(* PLC project AgentPLC, Beckhoff Automation GmbH TwinCAT PLC Control 3.5.21.61 *)
(* stored: creationDateTime 2026-11-03T10:24:45.563819, modificationDateTime 2026-11-03T10:24:45.5668157 *)

PROGRAM MAIN
VAR
	StartPB : BOOL;
	StopNC : BOOL;
	EStopHealthy : BOOL;
	PartSensor : BOOL;
	CountReset : BOOL;
	RunReq : BOOL;
	Horn : BOOL;
	Motor : BOOL;
	BatchLamp : BOOL;
	StartDelay : TON;
	BatchCounter : CTU;
END_VAR

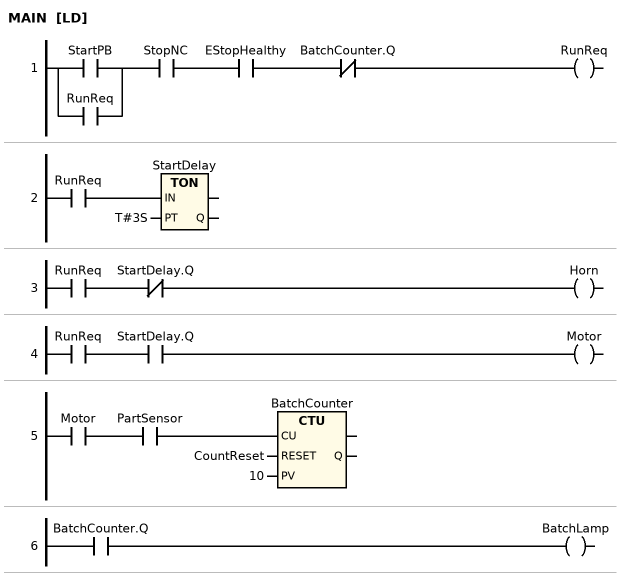
(* LD diagram, written out as Structured Text *)
(* Start/stop seal-in with E-stop permissive *)

RunReq := (StartPB OR RunReq) AND StopNC AND EStopHealthy AND NOT BatchCounter.Q;
(* Three-second start delay *)

StartDelay(IN := RunReq, PT := T#3S);
(* Horn during start delay *)

Horn := RunReq AND NOT StartDelay.Q;
(* Motor after start delay *)

Motor := RunReq AND StartDelay.Q;
(* Count ten parts; independent reset *)

BatchCounter(CU := Motor AND PartSensor, RESET := CountReset, PV := 10);
(* Batch-complete lamp *)

BatchLamp := BatchCounter.Q;
END_PROGRAM

CONFIGURATION Application
  RESOURCE AgentPLC ON PLC
    TASK PlcTask(INTERVAL := T#0ms, PRIORITY := 20);
    PROGRAM MAIN WITH PlcTask : MAIN;
  END_RESOURCE
END_CONFIGURATION
